(* IEC 61131-3 sources: PLC-Static-Analysis/modules/plc-rules/src/test/resources/PLCA-P005, 2 files *)

(* ---- compliant.st ---- *)
FUNCTION F_Safe : INT
VAR_INPUT
    pA : POINTER TO INT;
    pB : POINTER TO INT;
    pC : POINTER TO INT;
END_VAR
VAR
    n : INT;
    pLocal : POINTER TO INT;
END_VAR
IF pA <> 0 THEN
    F_Safe := pA^;
END_IF
IF pB = 0 THEN
    RETURN;
END_IF
F_Safe := F_Safe + pB^;
IF 0 <> pC AND_THEN pC^ > 0 THEN
    F_Safe := 1;
END_IF
pLocal := ADR(n);
F_Safe := F_Safe + pLocal^;
END_FUNCTION

(* ---- noncompliant.st ---- *)
FUNCTION F_Read : INT
VAR_INPUT
    pValue : POINTER TO INT;
    pOther : POINTER TO INT;
END_VAR
F_Read := pValue^; // PLCA-P005
F_Read := F_Read + pValue^;
IF F_Read > 0 THEN
    F_Read := pOther^; // PLCA-P005
END_IF
END_FUNCTION
